RESOURCE RES0 : EMB_RES_ECO
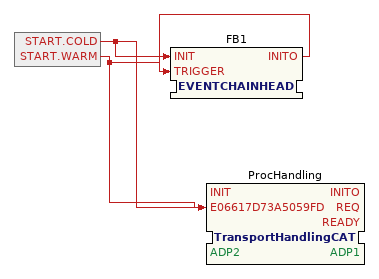
  FBS
    FB1 : EVENTCHAINHEAD;
    ProcHandling : TransportHandlingCAT;
  END_FBS
  EVENT_CONNECTIONS
    START.COLD TO FB1.INIT;
    START.WARM TO FB1.INIT;
    FB1.INITO TO FB1.TRIGGER;
    START.COLD TO ProcHandling.E06617D73A5059FD;
    START.WARM TO ProcHandling.E06617D73A5059FD;
  END_CONNECTIONS
END_RESOURCE
